FUNCTION_BLOCK FB_EvalSafeDevice
VAR_INPUT
	iDevice:structSafeInputDevice;
	iMsgMask:BOOL;
END_VAR
VAR_OUTPUT
	qDeviceActuated:BOOL;
	qReadyForReset:BOOL;
	qReadyForReIntag:BOOL;
	qDiscpFault:BOOL;
	qDeviceOK:BOOL;
END_VAR
VAR
	timCheckDiscp: TON;
	tDiscrapFault: BOOL;
END_VAR
VAR // added by the converter: edge detectors and wires of the graphical bodies
    _w1 : BOOL;
END_VAR

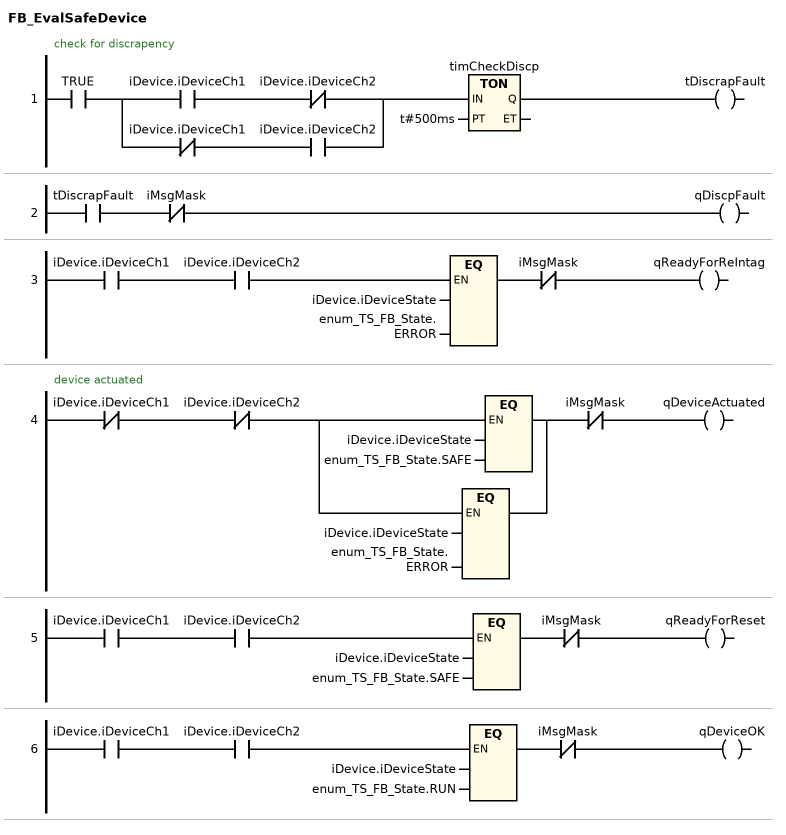
// NETWORK 1
// check for discrapency
timCheckDiscp(IN := TRUE AND (iDevice.iDeviceCh1 AND NOT iDevice.iDeviceCh2 OR NOT iDevice.iDeviceCh1 AND iDevice.iDeviceCh2), PT := t#500ms); // TON
tDiscrapFault := timCheckDiscp.Q;

// NETWORK 2
qDiscpFault := tDiscrapFault AND NOT iMsgMask;

// NETWORK 3
qReadyForReIntag := (iDevice.iDeviceCh1 AND iDevice.iDeviceCh2 AND iDevice.iDeviceState = enum_TS_FB_State.ERROR) AND NOT iMsgMask;

// NETWORK 4
// device actuated
_w1 := NOT iDevice.iDeviceCh1 AND NOT iDevice.iDeviceCh2;
qDeviceActuated := (_w1 AND iDevice.iDeviceState = enum_TS_FB_State.SAFE OR _w1 AND iDevice.iDeviceState = enum_TS_FB_State.ERROR) AND NOT iMsgMask;

// NETWORK 5
qReadyForReset := (iDevice.iDeviceCh1 AND iDevice.iDeviceCh2 AND iDevice.iDeviceState = enum_TS_FB_State.SAFE) AND NOT iMsgMask;

// NETWORK 6
qDeviceOK := (iDevice.iDeviceCh1 AND iDevice.iDeviceCh2 AND iDevice.iDeviceState = enum_TS_FB_State.RUN) AND NOT iMsgMask;

END_FUNCTION_BLOCK

(* stored: Version 1.1.0.1, ProductVersion 3.1.4024.11
   POU FB_EvalSafeDevice: Id {91d722c8-2db1-0b16-121d-27b566274a83}, SpecialFunc None *)
